(* IEC 61131-3 sources: plcassist-cli/packages/volt-lsp-iec/test-corpus/awa-palletizer/Device/Plc Logic/Application/Library Manager/IODrvEtherCAT, 61 files *)

(* ---- ETC_CONSTANTS.gvl ---- *)
VAR_GLOBAL
	_ETC_NUMBER_OF_MASTERS : INT := 1;
	_ETC_NUMBER_OF_SLAVES : INT := 1;
	_ETC_NUMBER_OF_SDO : INT := 0;
	_ETC_NUMBER_OF_INPUT_BYTES : INT := 0;
	_ETC_NUMBER_OF_OUTPUT_BYTES : INT := 0;
	_ETC_SYSTEM_HAS_INTEL_BYTEORDER : BOOL := TRUE;
END_VAR

(* ---- L_ETC_GLOBALS.gvl ---- *)
VAR_GLOBAL
	L_ETC_CMPID_IODRVETC : UDINT := 16#2006;
	L_ETC_EVT_PARAMETERTRANSFER_SERVICE : UDINT := 16#10000003;
END_VAR

(* ---- L_ETC_HC_GROUP_ITF.itf ---- *)
INTERFACE L_ETC_HC_GROUP_ITF
END_INTERFACE

(* ---- GETBOOLEANPROPERTY.fun ---- *)
FUNCTION GETBOOLEANPROPERTY : BOOL
VAR_INPUT
	STKEY : WSTRING;
END_VAR
END_FUNCTION

(* ---- GETCOMPANY.fun ---- *)
FUNCTION GETCOMPANY : WSTRING
END_FUNCTION

(* ---- GETNUMBERPROPERTY.fun ---- *)
FUNCTION GETNUMBERPROPERTY : DINT
VAR_INPUT
	STKEY : WSTRING;
END_VAR
END_FUNCTION

(* ---- GETTEXTPROPERTY.fun ---- *)
FUNCTION GETTEXTPROPERTY : WSTRING
VAR_INPUT
	STKEY : WSTRING;
END_VAR
END_FUNCTION

(* ---- GETTEXTPROPERTY2.fun ---- *)
FUNCTION GETTEXTPROPERTY2 : POINTER TO WSTRING
VAR_INPUT
	STKEY : WSTRING;
END_VAR
END_FUNCTION

(* ---- GETTITLE.fun ---- *)
FUNCTION GETTITLE : WSTRING
END_FUNCTION

(* ---- GETVERSION.fun ---- *)
FUNCTION GETVERSION : VERSION
END_FUNCTION

(* ---- GETVERSIONPROPERTY.fun ---- *)
FUNCTION GETVERSIONPROPERTY : VERSION
VAR_INPUT
	STKEY : WSTRING;
END_VAR
END_FUNCTION

(* ---- L_ETC_GETERRORSTRING.fun ---- *)
FUNCTION L_ETC_GETERRORSTRING : STRING(256)
VAR_INPUT
	EERRORCODE : L_ETC_ERRORCODE;
	ELANGUAGE : L_ETC_LANGUAGE := eng;
END_VAR
END_FUNCTION

(* ---- L_ETC_GETMASTER.fun ---- *)
FUNCTION L_ETC_GETMASTER : POINTER TO L_IODrvEtherCAT
VAR_INPUT
	USICOM : USINT;
END_VAR
END_FUNCTION

(* ---- L_ETC_GETSLAVE.fun ---- *)
FUNCTION L_ETC_GETSLAVE : POINTER TO ETCSlave
VAR_INPUT
	UIDEVICE : UINT;
END_VAR
END_FUNCTION

(* ---- L_ETC_HC_GETGROUP.fun ---- *)
FUNCTION L_ETC_HC_GETGROUP : L_ETC_HC_GROUP_ITF
VAR_INPUT
	USICOM : USINT := 1;
	GROUPNUMBER : UINT;
END_VAR
END_FUNCTION

(* ---- L_ETC_HC_GETGROUPCOUNT.fun ---- *)
FUNCTION L_ETC_HC_GETGROUPCOUNT : UINT
VAR_INPUT
	USICOM : USINT := 1;
END_VAR
END_FUNCTION

(* ---- L_ETC_HC_GETSLAVESOFGROUP.fun ---- *)
FUNCTION L_ETC_HC_GETSLAVESOFGROUP : DWORD
VAR_INPUT
	USICOM : USINT := 1;
	GROUPNUMBER : UINT;
	COUNT : POINTER TO UINT;
	SLAVES : POINTER TO POINTER TO ETCSlave;
END_VAR
END_FUNCTION

(* ---- L_ETC_IOCONTROL.fun ---- *)
FUNCTION L_ETC_IOCONTROL : DWORD
VAR_INPUT
	DWCODE : DWORD;
	PPARMS : POINTER TO L_ETC_IOCTLOPARMS;
END_VAR
END_FUNCTION

(* ---- ETCSLAVE.fb ---- *)
FUNCTION_BLOCK ETCSLAVE
VAR_INPUT
	XSETOPERATIONAL : BOOL;
END_VAR
VAR_OUTPUT
	XDONE : BOOL;
	XBUSY : BOOL;
	XERROR : BOOL;
	EERRORCODE : L_ETC_ERRORCODE;
	WSTATE : WORD;
END_VAR
VAR
	M_PIOCONFIGCONNECTOR : POINTER TO IoConfigConnector;
	M_SZPATH : STRING;
	M_SZNAME : STRING;
	M_DWVENDORID : DWORD;
	M_DWPRODUCTID : DWORD;
	M_DWREVISIONID : DWORD;
	M_UIPHYSSLAVEADDR : UINT;
	M_XDCENABLE : BOOL;
	M_XSETOPERATIONALLAST : BOOL;
	M_WSLAVESTATEACT : WORD;
	FBSLAVE2 : ETCSlave2;
	M_HCINIT : BOOL;
	M_HCINTERFACE : L_ETC_HC_GROUP_ITF;
	M_HCROLE : L_ETC_HC_ROLE;
	M_PMSSELECTIONPAR : POINTER TO IoStandard.IoConfigParameter;
	M_PMSSELECTION : USINT;
	MODULEHANDLERBASE : L_IMHP_ModuleHandler;
	M_SCOMMPATH : STRING(199);
	SLAVEADDRESS : UINT;
	REGISTERONCOMPONENTDIRECTORY : L_IC1P_RegisterOnComponentDirectory;
	M_ITFEVENTCALLBACK : CmpEventMgr.ICmpEventCallback;
	M_HEVENTUPDATECONFIGURATIONDONE : RTS_IEC_HANDLE;
	M_HINTERFACEUPDATECONFIGURATIONDONE : RTS_IEC_HANDLE;
	DCENABLE : BOOL;
	HCGROUP : L_ETC_HC_GROUP_ITF;
	HCROLE : L_ETC_HC_ROLE;
	IODRVETHERCAT : POINTER TO L_IODrvEtherCAT;
	ISMANDATORY : BOOL;
	ISPRESENT : BOOL;
	MODULEHANDLER : L_IMHP_IModuleHandler;
	NAME : STRING;
	PARAMETERSET : USINT;
	PHYSSLAVEADDR : UINT;
	WCSTATE : BOOL;
END_VAR
END_FUNCTION_BLOCK

METHOD EVENTCALLBACK : UDINT
VAR_INPUT
	PEVENTPARAM : POINTER TO EventParam;
END_VAR
END_METHOD

METHOD FB_EXIT : BOOL
VAR_INPUT
	BINCOPYCODE : BOOL;
END_VAR
END_METHOD

METHOD INITIALIZE : UDINT
VAR_INPUT
	WMODULETYPE : UINT;
	DWINSTANCE : UDINT;
	PCONNECTOR : POINTER TO IoConfigConnector;
END_VAR
END_METHOD

METHOD FB_INIT : BOOL
VAR_INPUT
	BINITRETAINS : BOOL;
	BINCOPYCODE : BOOL;
END_VAR
END_METHOD

(* ---- ETCSLAVE2.fb ---- *)
FUNCTION_BLOCK ETCSLAVE2
VAR_INPUT
	XSETOPERATIONAL : BOOL;
END_VAR
VAR_OUTPUT
	XDONE : BOOL;
	XBUSY : BOOL;
	XERROR : BOOL;
	EERRORCODE : L_ETC_ERRORCODE;
	WSTATE : WORD;
END_VAR
VAR
	M_PIOCONFIGCONNECTOR : POINTER TO IoConfigConnector;
	M_XSETOPERATIONALLAST : BOOL;
	M_UIPHYSSLAVEADDR : UINT;
	M_ADWJOBDATA : ARRAY [0..31] OF DWORD;
	GETSTATE : WORD;
	HCGROUP : L_ETC_HC_GROUP_ITF;
	HCROLE : L_ETC_HC_ROLE;
	IODRVETHERCAT : POINTER TO L_IODrvEtherCAT;
	ISMANDATORY : BOOL;
	PHYSSLAVEADDR : UINT;
END_VAR
END_FUNCTION_BLOCK

METHOD INITIALIZE : UDINT
VAR_INPUT
	WMODULETYPE : UINT;
	DWINSTANCE : UDINT;
	PCONNECTOR : POINTER TO IoConfigConnector;
END_VAR
END_METHOD

METHOD SETETCSLAVE
VAR_INPUT
	PCONNECTOR : POINTER TO IoConfigConnector;
	PETCSLAVE : POINTER TO ETCSlave;
END_VAR
END_METHOD

(* ---- ETCSLAVE_DIAG.fb ---- *)
FUNCTION_BLOCK ETCSLAVE_DIAG EXTENDS ETCSlave
VAR
	M_TREE : CAADiagTreeBase;
	CHILDNODECOUNT : CAA.COUNT;
	CONNECTOR : POINTER TO IoStandard.IoConfigConnector;
	ENABLE : BOOL;
	FIRSTCHILDNODE : DED.INode;
	INDEX : UDINT;
	ISROOTNODE : BOOL;
	NEXTSIBLINGNODE : DED.INode;
	PARENTNODE : DED.INode;
	SIBLINGNODECOUNT : CAA.COUNT;
END_VAR
END_FUNCTION_BLOCK

METHOD GETCHILD : DED.INode
VAR_INPUT
	UDIINDEX : UDINT;
END_VAR
END_METHOD

METHOD GETDEVICEDIAGNOSISINFO : DED.ERROR
VAR_INPUT
	PDATA : CAA.PVOID;
	SZSIZE : CAA.SIZE;
END_VAR
VAR_OUTPUT
	SZCOUNT : CAA.SIZE;
END_VAR
END_METHOD

METHOD GETDEVICEERRORASYNC : DED.PROC_STATE
VAR_INPUT
	ECMD : DED.PROC_CMD;
END_VAR
VAR_OUTPUT
	EERROR : DED.ERROR;
END_VAR
VAR_IN_OUT
	ERIDEVICEERROR : DED.ERROR_INFO;
END_VAR
END_METHOD

METHOD GETDEVICEINFO : DED.ERROR
VAR_IN_OUT
	DEIINFO : DED.DEVICE_INFO;
END_VAR
END_METHOD

METHOD GETDEVICESTATE : DED.DEVICE_STATE
VAR_OUTPUT
	XDIAGNOSISINFOAVAILABLE : BOOL;
	EERROR : DED.ERROR;
END_VAR
END_METHOD

METHOD GETSPECIFICDEVICEERRORASYNC : DED.PROC_STATE
VAR_INPUT
	ECMD : DED.PROC_CMD;
	PDATA : CAA.PVOID;
	SZSIZE : CAA.SIZE;
END_VAR
VAR_OUTPUT
	SZCOUNT : CAA.SIZE;
	EERROR : DED.ERROR;
END_VAR
END_METHOD

METHOD GETSPECIFICDEVICESTATE : DED.ERROR
VAR_INPUT
	PDATA : CAA.PVOID;
	SZSIZE : CAA.SIZE;
END_VAR
VAR_OUTPUT
	SZCOUNT : CAA.SIZE;
END_VAR
END_METHOD

METHOD INITIALIZE_DIAG : UDINT
VAR_INPUT
	PCONNECTOR : POINTER TO IoStandard.IoConfigConnector;
	NCONNECTORCOUNT : DINT;
	PARENT : POINTER TO DED.INode;
	CHILDREN : POINTER TO DED.INode;
	UDICHILDCOUNT : UDINT;
END_VAR
END_METHOD

METHOD SETCOMMUNICATIONSTATE : DED.ERROR
VAR_INPUT
	EREQUESTEDSTATE : DED.DEVICE_TRANSITION_STATE;
END_VAR
END_METHOD

(* ---- GLOBALTEXTLIST.fb ---- *)
FUNCTION_BLOCK GLOBALTEXTLIST
VAR
	M_TEXTLISTFILE : STRING(255);
	_STNAMESPACE : STRING;
END_VAR
END_FUNCTION_BLOCK

(* ---- L_ETC_CLEARCOUNTER.fb ---- *)
FUNCTION_BLOCK L_ETC_CLEARCOUNTER
VAR_INPUT
	XEXECUTE : BOOL;
	ECOUNTER : L_ETC_CLEARCOUNTER_COUNTER;
END_VAR
VAR_OUTPUT
	XDONE : BOOL;
	XBUSY : BOOL;
	XERROR : BOOL;
	EERRORCODE : L_ETC_ERRORCODE;
END_VAR
VAR
	XEXECUTELAST : BOOL;
	ADWJOBDATA : ARRAY [0..31] OF DWORD;
END_VAR
END_FUNCTION_BLOCK

(* ---- L_ETC_COE_SDOREAD.fb ---- *)
FUNCTION_BLOCK L_ETC_COE_SDOREAD
VAR_INPUT
	XEXECUTE : BOOL;
	XABORT : BOOL := FALSE;
	USICOM : USINT := 1;
	UIDEVICE : UINT;
	WINDEX : WORD;
	BYSUBINDEX : BYTE;
	UDITIMEOUT : UDINT;
	PBUFFER : CAA_PVOID := 0;
	SZSIZE : CAA_SIZE := 0;
END_VAR
VAR_OUTPUT
	XDONE : BOOL;
	XBUSY : BOOL;
	XERROR : BOOL;
	EERRORCODE : L_ETC_ERRORCODE;
	UDISDOABORT : UDINT;
	SZDATAREAD : CAA_SIZE;
END_VAR
VAR
	XEXECUTELAST : BOOL;
	ADWJOBDATA : ARRAY [0..31] OF DWORD;
END_VAR
END_FUNCTION_BLOCK

(* ---- L_ETC_COE_SDOREAD4.fb ---- *)
FUNCTION_BLOCK L_ETC_COE_SDOREAD4
VAR_INPUT
	XEXECUTE : BOOL;
	XABORT : BOOL := FALSE;
	USICOM : USINT := 1;
	UIDEVICE : UINT;
	WINDEX : WORD;
	BYSUBINDEX : BYTE;
	UDITIMEOUT : UDINT;
END_VAR
VAR_OUTPUT
	XDONE : BOOL;
	XBUSY : BOOL;
	XERROR : BOOL;
	EERRORCODE : L_ETC_ERRORCODE;
	UDISDOABORT : UDINT;
	ABYDATA : ARRAY [0..3] OF BYTE;
	SZDATAREAD : CAA_SIZE;
END_VAR
VAR
	SDOREAD : L_ETC_CoE_SdoRead;
END_VAR
END_FUNCTION_BLOCK

(* ---- L_ETC_COE_SDOREADEX.fb ---- *)
FUNCTION_BLOCK L_ETC_COE_SDOREADEX
VAR_INPUT
	XEXECUTE : BOOL;
	XABORT : BOOL := FALSE;
	USICOM : USINT := 1;
	UIDEVICE : UINT;
	DWFLAGS : DWORD;
	WINDEX : WORD;
	BYSUBINDEX : BYTE;
	UDITIMEOUT : UDINT;
	PBUFFER : CAA_PVOID := 0;
	SZSIZE : CAA_SIZE := 0;
END_VAR
VAR_OUTPUT
	XDONE : BOOL;
	XBUSY : BOOL;
	XERROR : BOOL;
	EERRORCODE : L_ETC_ERRORCODE;
	UDISDOABORT : UDINT;
	SZDATAREAD : CAA_SIZE;
END_VAR
VAR
	XEXECUTELAST : BOOL;
	ADWJOBDATA : ARRAY [0..31] OF DWORD;
END_VAR
END_FUNCTION_BLOCK

(* ---- L_ETC_COE_SDOWRITE.fb ---- *)
FUNCTION_BLOCK L_ETC_COE_SDOWRITE
VAR_INPUT
	XEXECUTE : BOOL;
	XABORT : BOOL := FALSE;
	USICOM : USINT := 1;
	UIDEVICE : UINT;
	WINDEX : WORD;
	BYSUBINDEX : BYTE;
	UDITIMEOUT : UDINT;
	PBUFFER : CAA_PVOID;
	SZSIZE : CAA_SIZE;
END_VAR
VAR_OUTPUT
	XDONE : BOOL;
	XBUSY : BOOL;
	XERROR : BOOL;
	EERRORCODE : L_ETC_ERRORCODE;
	UDISDOABORT : UDINT;
END_VAR
VAR
	XEXECUTELAST : BOOL;
	ADWJOBDATA : ARRAY [0..31] OF DWORD;
END_VAR
END_FUNCTION_BLOCK

(* ---- L_ETC_COE_SDOWRITE4.fb ---- *)
FUNCTION_BLOCK L_ETC_COE_SDOWRITE4
VAR_INPUT
	XEXECUTE : BOOL;
	XABORT : BOOL := FALSE;
	USICOM : USINT := 1;
	UIDEVICE : UINT;
	WINDEX : WORD;
	BYSUBINDEX : BYTE;
	UDITIMEOUT : UDINT;
	ABYDATA : ARRAY [0..3] OF BYTE;
	USIDATALENGTH : USINT;
END_VAR
VAR_OUTPUT
	XDONE : BOOL;
	XBUSY : BOOL;
	XERROR : BOOL;
	EERRORCODE : L_ETC_ERRORCODE;
	UDISDOABORT : UDINT;
END_VAR
VAR
	USILEN : USINT;
	SDOWRITE : L_ETC_CoE_SdoWrite;
END_VAR
END_FUNCTION_BLOCK

(* ---- L_ETC_COE_SDOWRITEEX.fb ---- *)
FUNCTION_BLOCK L_ETC_COE_SDOWRITEEX
VAR_INPUT
	XEXECUTE : BOOL;
	XABORT : BOOL := FALSE;
	USICOM : USINT := 1;
	UIDEVICE : UINT;
	DWFLAGS : DWORD;
	WINDEX : WORD;
	BYSUBINDEX : BYTE;
	UDITIMEOUT : UDINT;
	PBUFFER : CAA_PVOID;
	SZSIZE : CAA_SIZE;
END_VAR
VAR_OUTPUT
	XDONE : BOOL;
	XBUSY : BOOL;
	XERROR : BOOL;
	EERRORCODE : L_ETC_ERRORCODE;
	UDISDOABORT : UDINT;
END_VAR
VAR
	XEXECUTELAST : BOOL;
	ADWJOBDATA : ARRAY [0..31] OF DWORD;
END_VAR
END_FUNCTION_BLOCK

(* ---- L_ETC_ENGINEERINGMODE.fb ---- *)
FUNCTION_BLOCK L_ETC_ENGINEERINGMODE
VAR_INPUT
	USICOM : USINT := 1;
	XENABLE : BOOL;
END_VAR
VAR_OUTPUT
	XBUSY : BOOL;
	XACTIVE : BOOL;
	XERROR : BOOL;
	EERRORCODE : L_ETC_ERRORCODE;
	ESTATE : L_ETC_ENGMODE_STATE;
END_VAR
VAR
	USTEP : UINT := 0;
	XENABLEPRE : BOOL;
	CMD : L_ETC_CMD_T;
	RESULT : DWORD;
	SMSTATE : UDINT;
	FBMASTER : POINTER TO L_IODrvEtherCAT;
END_VAR
END_FUNCTION_BLOCK

(* ---- L_ETC_FOE_READ.fb ---- *)
FUNCTION_BLOCK L_ETC_FOE_READ
VAR_INPUT
	XEXECUTE : BOOL;
	XABORT : BOOL := FALSE;
	USICOM : USINT := 1;
	UIDEVICE : UINT;
	SFILENAME : CAA_FILENAME := '';
	SZFILENAMELEN : CAA_SIZE := 0;
	DWPASSWD : DWORD;
	UDITIMEOUT : UDINT;
	PBUFFER : CAA_PVOID := 0;
	SZSIZE : CAA_SIZE := 0;
END_VAR
VAR_OUTPUT
	XDONE : BOOL;
	XBUSY : BOOL;
	XERROR : BOOL;
	EERRORCODE : L_ETC_ERRORCODE;
	SZDATAREAD : CAA_SIZE;
END_VAR
VAR
	XEXECUTELAST : BOOL;
	ADWJOBDATA : ARRAY [0..31] OF DWORD;
END_VAR
END_FUNCTION_BLOCK

(* ---- L_ETC_FOE_WRITE.fb ---- *)
FUNCTION_BLOCK L_ETC_FOE_WRITE
VAR_INPUT
	XEXECUTE : BOOL;
	XABORT : BOOL := FALSE;
	USICOM : USINT := 1;
	UIDEVICE : UINT;
	SFILENAME : CAA_FILENAME := '';
	SZFILENAMELEN : CAA_SIZE := 0;
	DWPASSWD : DWORD;
	UDITIMEOUT : UDINT;
	PBUFFER : CAA_PVOID := 0;
	SZSIZE : CAA_SIZE := 0;
END_VAR
VAR_OUTPUT
	XDONE : BOOL;
	XBUSY : BOOL;
	XERROR : BOOL;
	EERRORCODE : L_ETC_ERRORCODE;
END_VAR
VAR
	XEXECUTELAST : BOOL;
	ADWJOBDATA : ARRAY [0..31] OF DWORD;
END_VAR
END_FUNCTION_BLOCK

(* ---- L_ETC_GETEMERGENCY.fb ---- *)
FUNCTION_BLOCK L_ETC_GETEMERGENCY
VAR_INPUT
	USICOM : USINT := 1;
	XEXECUTE : BOOL;
	XRESET : BOOL;
END_VAR
VAR_OUTPUT
	XDONE : BOOL;
	XBUSY : BOOL;
	XERROR : BOOL;
	EERRORCODE : L_ETC_ERRORCODE;
	OEMCY : L_ETC_COE_EMERGENCY;
	UICOUNT : UINT;
END_VAR
VAR
	M_XEXECUTELAST : BOOL;
	M_XRESETLAST : BOOL;
END_VAR
END_FUNCTION_BLOCK

METHOD DEINITIALIZE : BOOL
END_METHOD

METHOD FB_INIT : BOOL
VAR_INPUT
	BINITRETAINS : BOOL;
	BINCOPYCODE : BOOL;
END_VAR
END_METHOD

METHOD FB_EXIT : BOOL
VAR_INPUT
	BINCOPYCODE : BOOL;
END_VAR
END_METHOD

METHOD INITIALIZE : BOOL
END_METHOD

(* ---- L_ETC_GETMASTERDIAGNOSTIC.fb ---- *)
FUNCTION_BLOCK L_ETC_GETMASTERDIAGNOSTIC
VAR_INPUT
	XRESET : BOOL;
END_VAR
VAR_OUTPUT
	XDONE : BOOL;
	XBUSY : BOOL;
	XERROR : BOOL;
	EERRORCODE : L_ETC_ERRORCODE;
	ODIAGNOSTIC : L_ETC_DIAGNOSTIC;
END_VAR
VAR
	M_UDILASTMESSAGEID : UDINT;
	M_XRESETLAST : BOOL;
END_VAR
END_FUNCTION_BLOCK

(* ---- L_ETC_GETMASTERSTATE.fb ---- *)
FUNCTION_BLOCK L_ETC_GETMASTERSTATE
VAR_INPUT
	XEXECUTE : BOOL;
	UDITIMEOUT : UDINT;
END_VAR
VAR_OUTPUT
	XDONE : BOOL;
	XBUSY : BOOL;
	XERROR : BOOL;
	EERRORCODE : L_ETC_ERRORCODE;
	WSTATE : WORD;
END_VAR
VAR
	XEXECUTELAST : BOOL;
	ADWJOBDATA : ARRAY [0..31] OF DWORD;
END_VAR
END_FUNCTION_BLOCK

(* ---- L_ETC_GETSLAVESTATE.fb ---- *)
FUNCTION_BLOCK L_ETC_GETSLAVESTATE
VAR_INPUT
	XEXECUTE : BOOL;
	UIDEVICE : UINT;
	UDITIMEOUT : UDINT;
END_VAR
VAR_OUTPUT
	XDONE : BOOL;
	XBUSY : BOOL;
	XERROR : BOOL;
	EERRORCODE : L_ETC_ERRORCODE;
	WSTATE : WORD;
END_VAR
VAR
	XEXECUTELAST : BOOL;
	ADWJOBDATA : ARRAY [0..31] OF DWORD;
END_VAR
END_FUNCTION_BLOCK

METHOD FB_INIT : BOOL
VAR_INPUT
	BINITRETAINS : BOOL;
	BINCOPYCODE : BOOL;
END_VAR
END_METHOD

(* ---- L_ETC_HC_GROUP.fb ---- *)
FUNCTION_BLOCK L_ETC_HC_GROUP
VAR
	M_HDEVMANAGER : RTS_IEC_HANDLE;
	M_HINTERFACE : L_ETC_HC_GROUP_ITF;
	M_USICOM : USINT := 1;
	M_GROUPNUMBER : UINT;
	M_NAME : STRING;
	M_GROUPHEAD : POINTER TO ETCSlave;
	M_IDENTVALUE : UINT;
	M_SLAVECOUNT : UINT;
	M_SLAVES : POINTER TO ETCSlave;
	M_GROUPPRESENT : BOOL;
	M_GROUPSTATESUMMARY : WORD;
	M_WCSTATE : BOOL;
	M_RESERVE : ARRAY [0..15] OF ULINT;
	GETGROUPHEAD : POINTER TO ETCSlave;
	GETGROUPPRESENT : BOOL;
	GETGROUPSTATESUMMARY : L_ETC_HC_GROUPSTATESUMMARY;
	GETIDENTIFICATIONVALUE : UINT;
	GETNAME : STRING;
	GETSLAVECOUNT : UINT;
	GETSLAVES : POINTER TO ETCSlave;
	GROUPHEAD : POINTER TO ETCSlave;
	GROUPNUMBER : UINT;
	GROUPPRESENT : BOOL;
	GROUPSTATESUMMARY : WORD;
	IDENTIFICATIONVALUE : UINT;
	NAME : STRING;
	SLAVECOUNT : UINT;
	SLAVES : POINTER TO ETCSlave;
	WCSTATE : BOOL;
END_VAR
END_FUNCTION_BLOCK

METHOD FB_INIT : BOOL
VAR_INPUT
	BINITRETAINS : BOOL;
	BINCOPYCODE : BOOL;
END_VAR
END_METHOD

METHOD GETGROUPNUMBER : UINT
VAR_INPUT
	HINTERFACE : L_ETC_HC_GROUP_ITF;
END_VAR
END_METHOD

(* ---- L_ETC_HC_SETGROUPSTATE.fb ---- *)
FUNCTION_BLOCK L_ETC_HC_SETGROUPSTATE
VAR_INPUT
	USICOM : USINT := 1;
	XEXECUTE : BOOL;
	UIGROUP : UINT;
	WSTATE : WORD;
	UDITIMEOUT : UDINT;
END_VAR
VAR_OUTPUT
	XDONE : BOOL;
	XBUSY : BOOL;
	XERROR : BOOL;
	EERRORCODE : L_ETC_ERRORCODE;
END_VAR
VAR
	XEXECUTELAST : BOOL;
	ADWJOBDATA : ARRAY [0..31] OF DWORD;
END_VAR
END_FUNCTION_BLOCK

(* ---- L_ETC_HC_SETSLAVEPORTSTATE.fb ---- *)
FUNCTION_BLOCK L_ETC_HC_SETSLAVEPORTSTATE
VAR_INPUT
	USICOM : USINT := 1;
	XEXECUTE : BOOL;
	UIDEVICE : UINT;
	UIPORT : UINT;
	XCLOSE : BOOL;
	XFORCE : BOOL;
	UDITIMEOUT : UDINT;
END_VAR
VAR_OUTPUT
	XDONE : BOOL;
	XBUSY : BOOL;
	XERROR : BOOL;
	EERRORCODE : L_ETC_ERRORCODE;
END_VAR
VAR
	XEXECUTELAST : BOOL;
	ADWJOBDATA : ARRAY [0..16] OF DWORD;
END_VAR
END_FUNCTION_BLOCK

(* ---- L_ETC_MMCASSIGNADDRESS.fb ---- *)
FUNCTION_BLOCK L_ETC_MMCASSIGNADDRESS
VAR_INPUT
	XEXECUTE : BOOL;
	UIPOSITION : UINT;
	UIDEVICE : UINT;
END_VAR
VAR_OUTPUT
	XDONE : BOOL;
	XBUSY : BOOL;
	XERROR : BOOL;
	EERRORCODE : L_ETC_ERRORCODE;
END_VAR
VAR
	FBEEPROMWRITE : L_ETC_WriteEEPROM_intern;
END_VAR
END_FUNCTION_BLOCK

(* ---- L_ETC_MMCCONTROLLER.fb ---- *)
FUNCTION_BLOCK L_ETC_MMCCONTROLLER
VAR_INPUT
	XEXECUTE : BOOL;
	XABORT : BOOL;
	ESERVICE : L_ETC_MMCSERVICE;
	SZCONFIGURATION : STRING;
	XRESETTOPOLOGYCHANGEDCOUNTER : BOOL;
END_VAR
VAR_OUTPUT
	XDONE : BOOL;
	XBUSY : BOOL;
	XERROR : BOOL;
	EERRORCODE : L_ETC_MMCSERVICEERROR;
	XABORTED : BOOL;
	ESERVICESTATE : L_ETC_MMCSERVICESTATE;
	UDITOPOLOGYCHANGEDCOUNTER : UDINT;
END_VAR
VAR
	FBMMC : L_ETC_MMCController_intern;
	ACTUALCONFIGURATION : STRING;
	RUNNINGSERVICE : L_ETC_MMCSERVICE;
END_VAR
END_FUNCTION_BLOCK

METHOD FB_INIT : BOOL
VAR_INPUT
	BINITRETAINS : BOOL;
	BINCOPYCODE : BOOL;
END_VAR
END_METHOD

(* ---- L_ETC_MMCCONTROLLER_INTERN.fb ---- *)
FUNCTION_BLOCK L_ETC_MMCCONTROLLER_INTERN
VAR_INPUT
	XEXECUTE : BOOL;
	XABORT : BOOL;
	ESERVICE : L_ETC_MMCSERVICE;
	SZCONFIGURATION : STRING;
	XRESETTOPOLOGYCHANGEDCOUNTER : BOOL;
END_VAR
VAR_OUTPUT
	XDONE : BOOL;
	XBUSY : BOOL;
	XERROR : BOOL;
	EERRORCODE : L_ETC_MMCSERVICEERROR;
	XABORTED : BOOL;
	ESERVICESTATE : L_ETC_MMCSERVICESTATE;
	UDITOPOLOGYCHANGEDCOUNTER : UDINT;
END_VAR
VAR
	ESERVICEACT : L_ETC_MMCSERVICE;
	SZCONFIGURATIONACT : STRING;
	XEXECUTEPRE : BOOL;
	XABORTPRE : BOOL;
	XRESETTOPOLOGYCHANGEDCOUNTERPRE : BOOL;
	ADATA : ARRAY [0..31] OF DWORD;
END_VAR
END_FUNCTION_BLOCK

METHOD INITIALIZE
END_METHOD

(* ---- L_ETC_MMCCONTROLLERBUS.fb ---- *)
FUNCTION_BLOCK L_ETC_MMCCONTROLLERBUS
VAR_INPUT
	XEXECUTE : BOOL;
	XABORT : BOOL;
	SZCONFIGURATION : STRING;
	ESERVICE : L_ETC_MMCSERVICE;
	XRESETTOPOLOGYCHANGEDCOUNTER : BOOL;
END_VAR
VAR_OUTPUT
	XDONE : BOOL;
	XBUSY : BOOL;
	XERROR : BOOL;
	XABORTED : BOOL;
	EERRORCODE : L_ETC_MMCSERVICEERROR;
	ESERVICESTATE : L_ETC_MMCSERVICESTATE;
	UDITOPOLOGYCHANGEDCOUNTER : UDINT;
END_VAR
VAR
	FBMMC : L_ETC_MMCController;
	POMASTER : POINTER TO L_IODrvEtherCAT;
	STATE : INT;
	XEXECUTELAST : BOOL;
	XABORTLAST : BOOL;
	FBTIMEOUT : TON;
	XREADY : BOOL;
	ACTUALCONFIGURATION : STRING;
	RUNNINGSERVICE : L_ETC_MMCSERVICE;
END_VAR
END_FUNCTION_BLOCK

METHOD RESETOUTPUTS
END_METHOD

METHOD SETOUTPUTS
VAR_INPUT
	EERRORCODE2 : L_ETC_MMCSERVICEERROR;
END_VAR
END_METHOD

(* ---- L_ETC_MMCREADADDRESS.fb ---- *)
FUNCTION_BLOCK L_ETC_MMCREADADDRESS
VAR_INPUT
	XEXECUTE : BOOL;
	UIDEVICE : UINT;
	UDITIMEOUT : UDINT;
END_VAR
VAR_OUTPUT
	XDONE : BOOL;
	XBUSY : BOOL;
	XERROR : BOOL;
	EERRORCODE : L_ETC_ERRORCODE;
	UIDEVICESSA : UINT;
END_VAR
VAR
	FBEEPROMREAD : L_ETC_ReadEEPROM_intern;
END_VAR
END_FUNCTION_BLOCK

(* ---- L_ETC_READEEPROM_INTERN.fb ---- *)
FUNCTION_BLOCK L_ETC_READEEPROM_INTERN
VAR_INPUT
	XEXECUTE : BOOL;
	USICOM : USINT := 1;
	UIDEVICE : UINT;
	BAUTOINCADDR : BOOL := 0;
	UDITIMEOUT : UDINT;
	UIWORDADDRESS : UINT;
	PBUFFER : CAA_PVOID := 0;
	SZSIZE : CAA_SIZE := 0;
END_VAR
VAR_OUTPUT
	XDONE : BOOL;
	XBUSY : BOOL;
	XERROR : BOOL;
	EERRORCODE : L_ETC_ERRORCODE;
	SZDATAREAD : CAA_SIZE;
END_VAR
VAR
	XEXECUTELAST : BOOL;
	ADWJOBDATA : ARRAY [0..31] OF DWORD;
END_VAR
END_FUNCTION_BLOCK

(* ---- L_ETC_READERRCNT.fb ---- *)
FUNCTION_BLOCK L_ETC_READERRCNT
VAR_INPUT
	XEXECUTE : BOOL;
	UIDEVICE : UINT;
END_VAR
VAR_OUTPUT
	XDONE : BOOL;
	XBUSY : BOOL;
	XERROR : BOOL;
	EERRORCODE : L_ETC_ERRORCODE;
	REDERRCNT : L_ETC_SLAVE_PORTS;
	GREENERRCNT : L_ETC_SLAVE_PORTS;
END_VAR
VAR
	WINDEX : WORD;
	XEXCECUTEOLD : BOOL;
	WSTATE : WORD;
	GETSLAVESTATE : L_ETC_GetSlaveState;
	MYEC_T_IOCTLPARMS : L_ETC_IOCTLOPARMS;
	RESULT : DWORD;
	SDOREAD : L_ETC_CoE_SdoRead;
	WMYDATA : WORD;
	DWMYLENGTH : CAA_SIZE := 2;
	BYSUBCODEOFFSET : BYTE;
END_VAR
END_FUNCTION_BLOCK

(* ---- L_ETC_READERRCNT2.fb ---- *)
FUNCTION_BLOCK L_ETC_READERRCNT2
VAR_INPUT
	XEXECUTE : BOOL;
	UIDEVICE : UINT;
END_VAR
VAR_OUTPUT
	XDONE : BOOL;
	XBUSY : BOOL;
	XERROR : BOOL;
	EERRORCODE : L_ETC_ERRORCODE;
	REDERRCNT : L_ETC_SLAVE_PORTS2;
	GREENERRCNT : L_ETC_SLAVE_PORTS;
END_VAR
VAR
	WINDEX : WORD;
	XEXCECUTEOLD : BOOL;
	WSTATE : WORD;
	GETSLAVESTATE : L_ETC_GetSlaveState;
	MYEC_T_IOCTLPARMS : L_ETC_IOCTLOPARMS;
	RESULT : DWORD;
	SDOREAD : L_ETC_CoE_SdoReadEx;
	WMYDATA : WORD;
	DWMYLENGTH : CAA_SIZE := 2;
	BYSUBCODEOFFSET : BYTE;
	EC_SLAVE_BASE_ADDRESS : WORD := 1001;
	EC_IOCTL_FORCE_SLVSTAT_COLLECTION : DWORD := 44;
	EC_SLAVE_CONF_AND_INFO_OBJECT_0X3000 : WORD := 16#3000;
	EC_MOD_BASE_SUBIDX_RX_ERR_CNT_PORT0 : BYTE := 24;
END_VAR
END_FUNCTION_BLOCK

METHOD RESETOUTPUT
END_METHOD

(* ---- L_ETC_READERRCNTREAD.fb ---- *)
FUNCTION_BLOCK L_ETC_READERRCNTREAD
VAR_INPUT
	USICOM : USINT := 1;
	XEXECUTE : BOOL;
	UIDEVICE : UINT;
END_VAR
VAR_OUTPUT
	XDONE : BOOL;
	XBUSY : BOOL;
	XERROR : BOOL;
	EERRORCODE : L_ETC_ERRORCODE;
	RXERRORCNT : L_ETC_SLAVE_PORTS2;
	FWDRXERRORCNT : L_ETC_SLAVE_PORTS;
	PROCESSINGUNITERRORCNT : BYTE;
	PDIERRORCNT : BYTE;
	LOSTLINKCNT : L_ETC_SLAVE_PORTS;
END_VAR
VAR
	XEXCECUTEOLD : BOOL;
	WSTATE : WORD;
	PSLAVE : POINTER TO ETCSlave;
	DWSLAVEID : DWORD;
	SLAVEDESC : L_ETC_SLVSTATISTICS_DESC2_T;
	OIOCTLPARAMS : L_ETC_IOCTLOPARMS;
	RESULT : DWORD;
	DWREAD : DWORD;
	EC_IOCTL_GET_SLVSTATISTICS : DWORD := 45;
END_VAR
END_FUNCTION_BLOCK

METHOD RESETOUTPUT
END_METHOD

(* ---- L_ETC_READERRCNTUPDATE.fb ---- *)
FUNCTION_BLOCK L_ETC_READERRCNTUPDATE
VAR_INPUT
	USICOM : USINT := 1;
	XEXECUTE : BOOL;
END_VAR
VAR_OUTPUT
	XDONE : BOOL;
	XBUSY : BOOL;
	XERROR : BOOL;
	EERRORCODE : L_ETC_ERRORCODE;
END_VAR
VAR
	XEXCECUTEOLD : BOOL;
	WSTATE : WORD;
	PMASTER : POINTER TO L_IODrvEtherCAT;
	UDICYCLETIME : DWORD;
	OIOCTLRPARAMS : L_ETC_IOCTLOPARMS;
	RESULT : DWORD;
	TIMER : TON;
	TVAL : TIME;
	EC_IOCTL_FORCE_SLVSTAT_COLLECTION : DWORD := 44;
END_VAR
END_FUNCTION_BLOCK

METHOD RESETOUTPUTS
END_METHOD

(* ---- L_ETC_REGISTERREAD.fb ---- *)
FUNCTION_BLOCK L_ETC_REGISTERREAD
VAR_INPUT
	XEXECUTE : BOOL;
	XABORT : BOOL := FALSE;
	USICOM : USINT := 1;
	XAUTOINCADDR : BOOL := 0;
	UIDEVICE : UINT;
	WREGISTER : WORD;
	UDITIMEOUT : UDINT;
	PBUFFER : CAA_PVOID := 0;
	SZSIZE : CAA_SIZE := 0;
END_VAR
VAR_OUTPUT
	XDONE : BOOL;
	XBUSY : BOOL;
	XERROR : BOOL;
	EERRORCODE : L_ETC_ERRORCODE;
	SZDATAREAD : CAA_SIZE;
END_VAR
VAR
	XEXECUTELAST : BOOL;
	ADWJOBDATA : ARRAY [0..31] OF DWORD;
END_VAR
END_FUNCTION_BLOCK

(* ---- L_ETC_REGISTERWRITE.fb ---- *)
FUNCTION_BLOCK L_ETC_REGISTERWRITE
VAR_INPUT
	XEXECUTE : BOOL;
	XABORT : BOOL := FALSE;
	USICOM : USINT := 1;
	XAUTOINCADDR : BOOL := 0;
	UIDEVICE : UINT;
	WREGISTER : WORD;
	UDITIMEOUT : UDINT;
	PBUFFER : CAA_PVOID := 0;
	SZSIZE : CAA_SIZE := 0;
END_VAR
VAR_OUTPUT
	XDONE : BOOL;
	XBUSY : BOOL;
	XERROR : BOOL;
	EERRORCODE : L_ETC_ERRORCODE;
END_VAR
VAR
	XEXECUTELAST : BOOL;
	ADWJOBDATA : ARRAY [0..31] OF DWORD;
END_VAR
END_FUNCTION_BLOCK

(* ---- L_ETC_RESETERRCNT.fb ---- *)
FUNCTION_BLOCK L_ETC_RESETERRCNT
VAR_INPUT
	XEXECUTE : BOOL;
END_VAR
VAR_OUTPUT
	XDONE : BOOL;
	XBUSY : BOOL;
	XERROR : BOOL;
	EERRORCODE : L_ETC_ERRORCODE;
END_VAR
VAR
	XEXCECUTEOLD : BOOL := 0;
	WSTATE : WORD;
	GETMASTERSTATE : L_ETC_GetMasterState;
	MYEC_T_IOCTLPARMS : L_ETC_IOCTLOPARMS;
	RESULT : DWORD := 0;
END_VAR
END_FUNCTION_BLOCK

(* ---- L_ETC_SETMASTERSTATE.fb ---- *)
FUNCTION_BLOCK L_ETC_SETMASTERSTATE
VAR_INPUT
	XEXECUTE : BOOL;
	WSTATE : WORD;
	UDITIMEOUT : UDINT;
END_VAR
VAR_OUTPUT
	XDONE : BOOL;
	XBUSY : BOOL;
	XERROR : BOOL;
	EERRORCODE : L_ETC_ERRORCODE;
END_VAR
VAR
	XEXECUTELAST : BOOL;
	ADWJOBDATA : ARRAY [0..31] OF DWORD;
END_VAR
END_FUNCTION_BLOCK

(* ---- L_ETC_SETSLAVESTATE.fb ---- *)
FUNCTION_BLOCK L_ETC_SETSLAVESTATE
VAR_INPUT
	XEXECUTE : BOOL;
	UIDEVICE : UINT;
	WSTATE : WORD;
	UDITIMEOUT : UDINT;
END_VAR
VAR_OUTPUT
	XDONE : BOOL;
	XBUSY : BOOL;
	XERROR : BOOL;
	EERRORCODE : L_ETC_ERRORCODE;
END_VAR
VAR
	XEXECUTELAST : BOOL;
	ADWJOBDATA : ARRAY [0..31] OF DWORD;
END_VAR
END_FUNCTION_BLOCK

(* ---- L_ETC_SETSLAVESTATEFWDL.fb ---- *)
FUNCTION_BLOCK L_ETC_SETSLAVESTATEFWDL
VAR_INPUT
	XEXECUTE : BOOL;
	UIDEVICE : UINT;
	WSTATE : WORD;
	UDITIMEOUT : UDINT;
END_VAR
VAR_OUTPUT
	XDONE : BOOL;
	XBUSY : BOOL;
	XERROR : BOOL;
	EERRORCODE : L_ETC_ERRORCODE;
END_VAR
VAR
	XEXECUTELAST : BOOL;
	ADWJOBDATA : ARRAY [0..31] OF DWORD;
END_VAR
END_FUNCTION_BLOCK

(* ---- L_ETC_VOE_WRITEREAD_INTERN.fb ---- *)
FUNCTION_BLOCK L_ETC_VOE_WRITEREAD_INTERN
VAR_INPUT
	XEXECUTE : BOOL;
	USICOM : USINT := 1;
	UIDEVICE : UINT;
	UDITIMEOUT : UDINT;
	USICHANNEL : USINT;
	UDIVENDORID : UDINT;
	UIVENDORTYPE : UINT;
	PBUFFERWRITE : CAA_PVOID;
	SZSIZEWRITE : CAA_SIZE;
	PBUFFERREAD : CAA_PVOID;
	SZSIZEREAD : CAA_SIZE;
END_VAR
VAR_OUTPUT
	XDONE : BOOL;
	XBUSY : BOOL;
	XERROR : BOOL;
	EERRORCODE : L_ETC_ERRORCODE;
	SZDATAREAD : CAA_SIZE;
END_VAR
VAR
	XEXECUTELAST : BOOL;
	ADWJOBDATA : ARRAY [0..31] OF DWORD;
END_VAR
END_FUNCTION_BLOCK

(* ---- L_ETC_WRITEEEPROM_INTERN.fb ---- *)
FUNCTION_BLOCK L_ETC_WRITEEEPROM_INTERN
VAR_INPUT
	XEXECUTE : BOOL;
	USICOM : USINT := 1;
	UIDEVICE : UINT;
	BAUTOINCADDR : BOOL := 0;
	UDITIMEOUT : UDINT;
	UIWORDADDRESS : UINT;
	PBUFFER : CAA_PVOID := 0;
	SZSIZE : CAA_SIZE := 0;
END_VAR
VAR_OUTPUT
	XDONE : BOOL;
	XBUSY : BOOL;
	XERROR : BOOL;
	EERRORCODE : L_ETC_ERRORCODE;
END_VAR
VAR
	XEXECUTELAST : BOOL;
	ADWJOBDATA : ARRAY [0..31] OF DWORD;
END_VAR
END_FUNCTION_BLOCK

(* ---- L_IODRVETHERCAT.fb ---- *)
FUNCTION_BLOCK L_IODRVETHERCAT
VAR_INPUT
	XRESTART : BOOL := FALSE;
	XSTOPBUS : BOOL := FALSE;
	XWAITWHILEBOOTINGCONTINUE : BOOL;
END_VAR
VAR_OUTPUT
	XDONE : BOOL;
	XBUSY : BOOL;
	XERROR : BOOL;
	EERRORCODE : L_ETC_ERRORCODE;
	WSTATE : WORD;
	XDISTRIBUTEDCLOCKINSYNC : BOOL;
	XWAITWHILEBOOTING : BOOL;
END_VAR
VAR
	M_PIOCONFIGCONNECTOR : POINTER TO IoConfigConnector;
	M_FBIODRVETHERCAT : L_IODrvEtherCAT_intern2;
	M_UDICYCLETIME : UDINT;
	M_NUMBEROFSLAVESCONFIGURED : UINT;
	M_IDX_NEXT : UINT;
	M_IDX_CHUNK : UINT := 3;
	MODULEHANDLERBASE : L_IMHP_ModuleHandler;
	CYCLETIME : UDINT;
	GETCONNECTOR : POINTER TO IoConfigConnector;
	MODULEHANDLER : L_IMHP_IModuleHandler;
	NUMBEROFSLAVESCONFIGURED : UINT;
	WCSTATE : BOOL;
END_VAR
END_FUNCTION_BLOCK

METHOD BEFOREREADINPUTS
END_METHOD

METHOD INITIALIZE : UDINT
VAR_INPUT
	WMODULETYPE : UINT;
	DWINSTANCE : UDINT;
	PCONNECTOR : POINTER TO IoConfigConnector;
END_VAR
END_METHOD

METHOD FB_INIT : BOOL
VAR_INPUT
	BINITRETAINS : BOOL;
	BINCOPYCODE : BOOL;
END_VAR
END_METHOD

(* ---- L_IODRVETHERCAT_DIAG.fb ---- *)
FUNCTION_BLOCK L_IODRVETHERCAT_DIAG EXTENDS L_IODrvEtherCAT
VAR
	M_TREE : CAADiagTreeBase;
	M_DIAG : L_ETC_GetMasterDiagnostic;
	CHILDNODECOUNT : CAA.COUNT;
	CONNECTOR : POINTER TO IoStandard.IoConfigConnector;
	ENABLE : BOOL;
	FIRSTCHILDNODE : DED.INode;
	INDEX : UDINT;
	ISROOTNODE : BOOL;
	NEXTSIBLINGNODE : DED.INode;
	PARENTNODE : DED.INode;
	SIBLINGNODECOUNT : CAA.COUNT;
END_VAR
END_FUNCTION_BLOCK

METHOD GETBUSDIAGNOSISINFO : DED.ERROR
VAR_INPUT
	PDATA : CAA.PVOID;
	SZSIZE : CAA.SIZE;
END_VAR
VAR_OUTPUT
	SZCOUNT : CAA.SIZE;
END_VAR
END_METHOD

METHOD GETBUSERRORASYNC : DED.PROC_STATE
VAR_INPUT
	ECMD : DED.PROC_CMD;
END_VAR
VAR_OUTPUT
	EERROR : DED.ERROR;
END_VAR
VAR_IN_OUT
	ERIBUSERROR : DED.ERROR_INFO;
END_VAR
END_METHOD

METHOD GETBUSINFO : DED.ERROR
VAR_IN_OUT
	BUIINFO : DED.BUS_INFO;
END_VAR
END_METHOD

METHOD GETBUSSTATE : DED.BUS_STATE
VAR_OUTPUT
	XDIAGNOSISINFOAVAILABLE : BOOL;
	EERROR : DED.ERROR;
END_VAR
END_METHOD

METHOD GETCHILD : DED.INode
VAR_INPUT
	UDIINDEX : UDINT;
END_VAR
END_METHOD

METHOD GETDEVICEDIAGNOSISINFO : DED.ERROR
VAR_INPUT
	PDATA : CAA.PVOID;
	SZSIZE : CAA.SIZE;
END_VAR
VAR_OUTPUT
	SZCOUNT : CAA.SIZE;
END_VAR
END_METHOD

METHOD GETDEVICEERRORASYNC : DED.PROC_STATE
VAR_INPUT
	ECMD : DED.PROC_CMD;
END_VAR
VAR_OUTPUT
	EERROR : DED.ERROR;
END_VAR
VAR_IN_OUT
	ERIDEVICEERROR : DED.ERROR_INFO;
END_VAR
END_METHOD

METHOD GETDEVICEINFO : DED.ERROR
VAR_IN_OUT
	DEIINFO : DED.DEVICE_INFO;
END_VAR
END_METHOD

METHOD GETDEVICESTATE : DED.DEVICE_STATE
VAR_OUTPUT
	XDIAGNOSISINFOAVAILABLE : BOOL;
	EERROR : DED.ERROR;
END_VAR
END_METHOD

METHOD GETQOS : DED.ERROR
VAR_IN_OUT
	QUALITYINFO : DED.QOS_INFO;
END_VAR
END_METHOD

METHOD GETSPECIFICBUSSTATE : DED.ERROR
VAR_INPUT
	PDATA : CAA.PVOID;
	SZSIZE : CAA.SIZE;
END_VAR
VAR_OUTPUT
	SZCOUNT : CAA.SIZE;
END_VAR
END_METHOD

METHOD GETSPECIFICDEVICEERRORASYNC : DED.PROC_STATE
VAR_INPUT
	ECMD : DED.PROC_CMD;
	PDATA : CAA.PVOID;
	SZSIZE : CAA.SIZE;
END_VAR
VAR_OUTPUT
	SZCOUNT : CAA.SIZE;
	EERROR : DED.ERROR;
END_VAR
END_METHOD

METHOD GETSPECIFICDEVICESTATE : DED.ERROR
VAR_INPUT
	PDATA : CAA.PVOID;
	SZSIZE : CAA.SIZE;
END_VAR
VAR_OUTPUT
	SZCOUNT : CAA.SIZE;
END_VAR
END_METHOD

METHOD INITIALIZE_DIAG : UDINT
VAR_INPUT
	PCONNECTOR : POINTER TO IoStandard.IoConfigConnector;
	NCONNECTORCOUNT : DINT;
	PARENT : POINTER TO DED.INode;
	CHILDREN : POINTER TO DED.INode;
	UDICHILDCOUNT : UDINT;
END_VAR
END_METHOD

METHOD SETCOMMUNICATIONSTATE : DED.ERROR
VAR_INPUT
	EREQUESTEDSTATE : DED.DEVICE_TRANSITION_STATE;
END_VAR
END_METHOD

(* ---- L_IODRVETHERCAT_INTERN.fb ---- *)
FUNCTION_BLOCK L_IODRVETHERCAT_INTERN
VAR_INPUT
	XRESTART : BOOL := FALSE;
	XSTOPBUS : BOOL := FALSE;
END_VAR
VAR_OUTPUT
	XDONE : BOOL;
	XBUSY : BOOL;
	XERROR : BOOL;
	EERRORCODE : L_ETC_ERRORCODE;
	WSTATE : WORD;
	XDISTRIBUTEDCLOCKINSYNC : BOOL;
END_VAR
VAR
	M_PIOCONFIGCONNECTOR : POINTER TO IoConfigConnector;
	M_WCOMMAND : UDINT;
	M_UDISTOPTIMEOUT : UDINT := 5000;
	M_UDISTARTTIMEOUT : UDINT := 60000;
	M_UDILASTMESSAGEID : UDINT;
	M_SLASTMESSAGE : STRING;
	M_WSTATEREQ : UINT;
	M_ADWJOBDATA : ARRAY [0..31] OF DWORD;
	M_XRESTARTLAST : BOOL;
	M_XSTOPBUSLAST : BOOL;
	NUMBEROFSLAVESCONFIGURED : UINT;
	WCSTATE : BOOL;
END_VAR
END_FUNCTION_BLOCK

METHOD BEFOREREADINPUTS
END_METHOD

METHOD INITIALIZE : UDINT
VAR_INPUT
	WMODULETYPE : UINT;
	DWINSTANCE : UDINT;
	PCONNECTOR : POINTER TO IoConfigConnector;
	PPARENT : POINTER TO L_IODrvEtherCAT;
END_VAR
END_METHOD

(* ---- L_IODRVETHERCAT_INTERN2.fb ---- *)
FUNCTION_BLOCK L_IODRVETHERCAT_INTERN2
VAR_INPUT
	XRESTART : BOOL := FALSE;
	XSTOPBUS : BOOL := FALSE;
	XWAITWHILEBOOTINGCONTINUE : BOOL;
	DWRESERVEINPUT : ARRAY [0..15] OF DWORD;
END_VAR
VAR_OUTPUT
	XDONE : BOOL;
	XBUSY : BOOL;
	XERROR : BOOL;
	EERRORCODE : L_ETC_ERRORCODE;
	WSTATE : WORD;
	XDISTRIBUTEDCLOCKINSYNC : BOOL;
	XWAITWHILEBOOTING : BOOL;
	DWRESERVEOUTPUT : ARRAY [0..15] OF DWORD;
END_VAR
VAR
	M_PIOCONFIGCONNECTOR : POINTER TO IoConfigConnector;
	M_WCOMMAND : UDINT;
	M_UDISTOPTIMEOUT : UDINT := 5000;
	M_UDISTARTTIMEOUT : UDINT := 60000;
	M_UDILASTMESSAGEID : UDINT;
	M_SLASTMESSAGE : STRING;
	M_WSTATEREQ : UINT;
	M_ADWJOBDATA : ARRAY [0..31] OF DWORD;
	M_XRESTARTLAST : BOOL;
	M_XSTOPBUSLAST : BOOL;
	DWRESERVEMEM : ARRAY [0..15] OF DWORD;
	NUMBEROFSLAVESCONFIGURED : UINT;
	WCSTATE : BOOL;
END_VAR
END_FUNCTION_BLOCK

METHOD BEFOREREADINPUTS
END_METHOD

METHOD INITIALIZE : UDINT
VAR_INPUT
	WMODULETYPE : UINT;
	DWINSTANCE : UDINT;
	PCONNECTOR : POINTER TO IoConfigConnector;
	PPARENT : POINTER TO L_IODrvEtherCAT;
END_VAR
END_METHOD
